Fanuc KAREL source: KB00115.KL

PROGRAM KB00115
%NOLOCKGROUP
%ENVIRONMENT KCLOP
VAR
BEGIN
  KCL_STATUS
END KB00115
